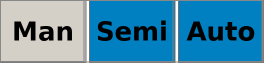
VISUALIZATION Mode_Select  // 264x63
VAR_IN_OUT
	stMode: ST_Mode;
END_VAR
    Button (0,0 86x63), "Man", colour toggle: stModeMain.iActMode=eManualMode
        OnMouseDown: execute {
            stModeMain.bSetManual:=TRUE;
            stMode.bSetSemi:=FALSE;
            stMode.bSetAuto:=FALSE;
        }
    Button (89,0 86x63), "Semi", colour toggle: stModeMain.iActMode=eSemiAutoMode
        OnMouseDown: execute {
            stModeMain.bSetManual:=FALSE;
            stMode.bSetSemi:=TRUE;
            stMode.bSetAuto:=FALSE;
        }
    Button (178,0 86x63), "Auto", colour toggle: stModeMain.iActMode=eAutoMode
        OnMouseDown: execute {
            stModeMain.bSetManual:=FALSE;
            stMode.bSetSemi:=FALSE;
            stMode.bSetAuto:=TRUE;
        }
END_VISUALIZATION

(* stored: Version 1.1.0.1, ProductVersion 3.1.4024.13
   Visu Mode_Select: Id {7cc5a97b-2a07-4618-9cfd-a15c268a44e1} *)
